// TIA Portal project "BlinkGemma" (V18)

(* hardware
DEVICE "S71500/ET200MP station_1"  S7-1500 station
   slot 0: "Telaio di montaggio_0"  Rack  6ES7 590-1***0-0AA0
   slot 1: "PLC_1"  CPU 1516-3 PN/DP  6ES7 516-3AN01-0AB0  V1.8
      slot 3: "Display CPU_1"  6ES7591-1BA00-0AA0
   slot 2: "DI 32x24VDC HF_1"  DI 32x24VDC HF  6ES7 521-1BL00-0AB0  V1.0
   slot 3: "DQ 32x24VDC/0.5A HF_1"  DQ 32x24VDC/0.5A HF  6ES7 522-1BL01-0AB0  V1.0
   slot 4: "AI 8xU/I/RTD/TC ST_1"  AI 8xU/I/RTD/TC ST  6ES7 531-7KF00-0AB0  V1.0
   slot 5: "AQ 4xU/I ST_1"  AQ 4xU/I ST  6ES7 532-5HD00-0AB0  V1.0
*)

// ===== PLC "PLC_1"  CPU 1516-3 PN/DP =====

VAR_GLOBAL   // PLC tag table "Tabella delle variabili standard"
   "bLamp" AT %M0.1 : Bool;
   "tmp" AT %M0.0 : Bool;
   "oLed" AT %Q0.0 : Bool;
END_VAR

DATA_BLOCK "DB1-GestioneTappe"   // DB2
{ S7_Optimized_Access := 'TRUE' }
VERSION : 0.1
   VAR
      Gemma : Array[0..15] of Bool;
      M1P : Array[0..15] of Bool;
   END_VAR
BEGIN
   // Gemma[0] : Gemma tappa 0
   // Gemma[1] : Gemma tappa 1
   // Gemma[2] : Gemma tappa 2
   // Gemma[3] : Gemma tappa 3
   // Gemma[4] : Gemma tappa 4
   // Gemma[5] : Gemma tappa 5
   // Gemma[6] : Gemma tappa 6
   // Gemma[7] : Gemma tappa 7
   // Gemma[8] : Gemma tappa 8
   // Gemma[9] : Gemma tappa 9
   // Gemma[10] : Gemma tappa 10
   // Gemma[11] : Gemma tappa 11
   // Gemma[12] : Gemma tappa 12
   // Gemma[13] : Gemma tappa 13
   // Gemma[14] : Gemma tappa 14
   // Gemma[15] : Gemma tappa 15
   // M1P[0] : Macchina 1 tappa 0
   // M1P[1] : Macchina 1 tappa 1
   // M1P[2] : Macchina 1 tappa 2
   // M1P[3] : Macchina 1 tappa 3
   // M1P[4] : Macchina 1 tappa 4
   // M1P[5] : Macchina 1 tappa 5
   // M1P[6] : Macchina 1 tappa 6
   // M1P[7] : Macchina 1 tappa 7
   // M1P[8] : Macchina 1 tappa 8
   // M1P[9] : Macchina 1 tappa 9
   // M1P[10] : Macchina 1 tappa 10
   // M1P[11] : Macchina 1 tappa 11
   // M1P[12] : Macchina 1 tappa 12
   // M1P[13] : Macchina 1 tappa 13
   // M1P[14] : Macchina 1 tappa 14
   // M1P[15] : Macchina 1 tappa 15
END_DATA_BLOCK

DATA_BLOCK "DB2-GestioneComandi"   // DB3
{ S7_Optimized_Access := 'TRUE' }
VERSION : 0.1
   VAR
      bAuto : Bool;   // Comando Automatico
      bMan : Bool;   // Comando Manuale
      bStop : Bool;   // Comando Stop
      bReset : Bool;   // Comando Reset
      bEmergenza : Bool;   // Comando EMERGENZA
      bLedManuale : Bool;   // Comando Led Manuale
   END_VAR
BEGIN
END_DATA_BLOCK

DATA_BLOCK "DB3-GestioneStati"   // DB4
{ S7_Optimized_Access := 'TRUE' }
VERSION : 0.1
   VAR
      sStop : Bool;   // Stato Stop
      sAuto : Bool;   // Stato Automatico
      sMan : Bool;   // Stato Manuale
      sAttesaStop : Bool;   // Stato Attesa Stop
   END_VAR
BEGIN
END_DATA_BLOCK

DATA_BLOCK "DB4-GestioneMacchine"   // DB5
{ S7_Optimized_Access := 'TRUE' }
VERSION : 0.1
   VAR
      bIni : Bool;   // Inizializzazione M1
      bRip : Bool;   // Macchina a riposo
      attEmergenza : Bool;   // Emergenza ATTIVATA
   END_VAR
BEGIN
END_DATA_BLOCK

// folder: System blocks/Program resources

DATA_BLOCK "IEC_Timer_0_DB"   // DB1
{ S7_Optimized_Access := 'TRUE' }
AUTHOR : Simatic
FAMILY : IEC
NAME : IEC_TMR
VERSION : 1.0
// stored: InstanceOfName IEC_TIMER
"IEC_TIMER"
BEGIN
END_DATA_BLOCK

// folder: (top level)

FUNCTION "FC1-BaseTempi" : Void   // FC1, LAD
{ S7_Optimized_Access := 'TRUE' }
VERSION : 0.1
   VAR_TEMP   // added for the SCL form of the ladder/FBD networks
      _w1 : Bool;
   END_VAR
BEGIN

REGION Network 1
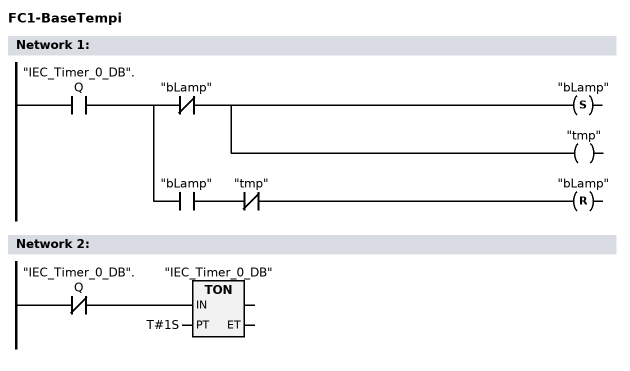
   RUNG wire#powerrail
      Contact( "IEC_Timer_0_DB".Q )
      wire#w1
      I_Contact( "bLamp" )
      wire#w2
      S_Coil( "bLamp" )
   END_RUNG
   RUNG wire#w2
      Coil( "tmp" )
   END_RUNG
   RUNG wire#w1
      Contact( "bLamp" )
      I_Contact( "tmp" )
      R_Coil( "bLamp" )
   END_RUNG
   // the same network as SCL:
   #_w1 := "IEC_Timer_0_DB".Q AND NOT "bLamp";
   IF #_w1 THEN "bLamp" := TRUE; END_IF;
   "tmp" := #_w1;
   IF "IEC_Timer_0_DB".Q AND "bLamp" AND NOT "tmp" THEN "bLamp" := FALSE; END_IF;
END_REGION

REGION Network 2
   "IEC_Timer_0_DB".TON(IN := NOT "IEC_Timer_0_DB".Q, PT := T#1S);
END_REGION
END_FUNCTION

FUNCTION "FC-Uscite" : Void   // FC2, LAD
{ S7_Optimized_Access := 'TRUE' }
VERSION : 0.1
BEGIN

REGION Network 1
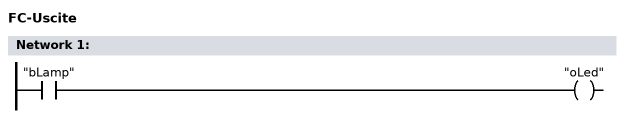
   RUNG wire#powerrail
      Contact( "bLamp" )
      Coil( "oLed" )
   END_RUNG
   // the same network as SCL:
   "oLed" := "bLamp";
END_REGION
END_FUNCTION

FUNCTION "FC3-GestioneGemma" : Void   // FC3, LAD
{ S7_Optimized_Access := 'TRUE' }
VERSION : 0.1
   VAR_TEMP   // added for the SCL form of the ladder/FBD networks
      _w1 : Bool;
      _w2 : Bool;
   END_VAR
BEGIN

REGION Network 1: Gestione: Tappa0 RESET Tappa0 e SET Tappa1 - oppure RESET Tappa0 SET Tappa3
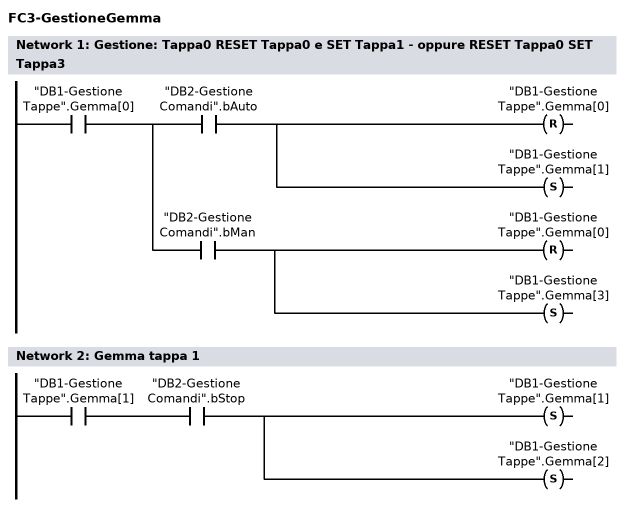
   RUNG wire#powerrail
      Contact( "DB1-GestioneTappe".Gemma[0] )
      wire#w1
      Contact( "DB2-GestioneComandi".bAuto )
      wire#w2
      R_Coil( "DB1-GestioneTappe".Gemma[0] )
   END_RUNG
   RUNG wire#w2
      S_Coil( "DB1-GestioneTappe".Gemma[1] )
   END_RUNG
   RUNG wire#w1
      Contact( "DB2-GestioneComandi".bMan )
      wire#w3
      R_Coil( "DB1-GestioneTappe".Gemma[0] )
   END_RUNG
   RUNG wire#w3
      S_Coil( "DB1-GestioneTappe".Gemma[3] )
   END_RUNG
   // the same network as SCL:
   #_w1 := "DB1-GestioneTappe".Gemma[0];
   #_w2 := "DB1-GestioneTappe".Gemma[0] AND "DB2-GestioneComandi".bAuto;
   IF #_w2 THEN
       "DB1-GestioneTappe".Gemma[0] := FALSE;
       "DB1-GestioneTappe".Gemma[1] := TRUE;
   END_IF;
   IF #_w1 AND "DB2-GestioneComandi".bMan THEN
       "DB1-GestioneTappe".Gemma[0] := FALSE;
       "DB1-GestioneTappe".Gemma[3] := TRUE;
   END_IF;
END_REGION

REGION Network 2: Gemma tappa 1
   RUNG wire#powerrail
      Contact( "DB1-GestioneTappe".Gemma[1] )
      Contact( "DB2-GestioneComandi".bStop )
      wire#w1
      S_Coil( "DB1-GestioneTappe".Gemma[1] )
   END_RUNG
   RUNG wire#w1
      S_Coil( "DB1-GestioneTappe".Gemma[2] )
   END_RUNG
   // the same network as SCL:
   #_w1 := "DB1-GestioneTappe".Gemma[1] AND "DB2-GestioneComandi".bStop;
   IF #_w1 THEN
       "DB1-GestioneTappe".Gemma[1] := TRUE;
       "DB1-GestioneTappe".Gemma[2] := TRUE;
   END_IF;
END_REGION
END_FUNCTION

FUNCTION "FC4-ResetPulsanti" : Void   // FC4, LAD
{ S7_Optimized_Access := 'TRUE' }
VERSION : 0.1
BEGIN

REGION Network 1: Reset Pulsante di STOP
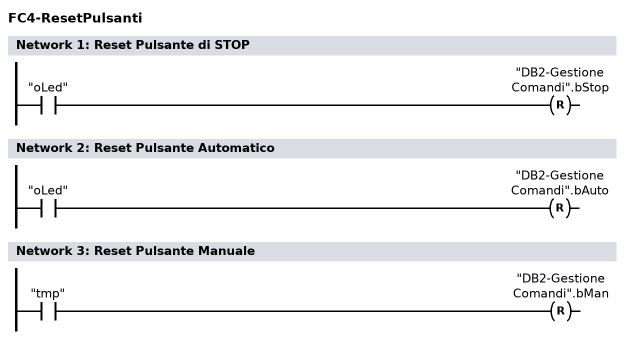
   RUNG wire#powerrail
      Contact( "oLed" )
      R_Coil( "DB2-GestioneComandi".bStop )
   END_RUNG
   // the same network as SCL:
   IF "oLed" THEN "DB2-GestioneComandi".bStop := FALSE; END_IF;
END_REGION

REGION Network 2: Reset Pulsante Automatico
   RUNG wire#powerrail
      Contact( "oLed" )
      R_Coil( "DB2-GestioneComandi".bAuto )
   END_RUNG
   // the same network as SCL:
   IF "oLed" THEN "DB2-GestioneComandi".bAuto := FALSE; END_IF;
END_REGION

REGION Network 3: Reset Pulsante Manuale
   RUNG wire#powerrail
      Contact( "tmp" )
      R_Coil( "DB2-GestioneComandi".bMan )
   END_RUNG
   // the same network as SCL:
   IF "tmp" THEN "DB2-GestioneComandi".bMan := FALSE; END_IF;
END_REGION
END_FUNCTION

ORGANIZATION_BLOCK "Main"   // OB1, LAD, ProgramCycle
TITLE = "Main Program Sweep (Cycle)"
{ S7_Optimized_Access := 'TRUE' }
VERSION : 0.1
   VAR_INPUT
      Initial_Call : Bool;   // Initial call of this OB
      Remanence : Bool;   // =True, if remanent data are available
   END_VAR
BEGIN

REGION Network 1
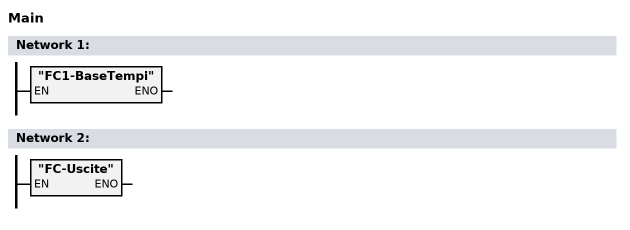
   RUNG wire#powerrail
      "FC1-BaseTempi"()
   END_RUNG
   // the same network as SCL:
   "FC1-BaseTempi"();
END_REGION

REGION Network 2
   RUNG wire#powerrail
      "FC-Uscite"()
   END_RUNG
   // the same network as SCL:
   "FC-Uscite"();
END_REGION
END_ORGANIZATION_BLOCK